// TIA Portal V21 export
// export: Created 2026-11-07T14:35:58.9708753Z, ExportSetting WithDefaults, DisplayName Totally Integrated Automation Portal, DisplayVersion V21, DisplayName STEP 7 Professional, DisplayVersion V21, DisplayName STEP 7 Safety, DisplayVersion V21, DisplayName Tech WebApplication, DisplayVersion V21, DisplayName WinCC Basic/Comfort/Advanced, DisplayVersion V21, DisplayName WinCC Unified, DisplayVersion V21
Screen "T07_Sym"  1024x768, Number=27
  ScreenLayer 
    SymbolicIOField "P_SymIO" at 0,0 size 100x30  CountVisibleItems=3, Mode=Output, OnValue=1, StyleItem=Symbolic I/O field, TextList=TL_State, TextOff="0", TextOn="1"
      ProcessValue := State
